// TIA Portal V21 export
// export: Created 2026-08-21T20:18:56.6399431Z, ExportSetting None, DisplayName Totally Integrated Automation Portal, DisplayVersion V21, DisplayName STEP 7 Professional, DisplayVersion V21, DisplayName STEP 7 Safety, DisplayVersion V21, DisplayName Tech WebApplication, DisplayVersion V21, DisplayName WinCC Basic/Comfort/Advanced, DisplayVersion V21, DisplayName WinCC Professional, DisplayVersion V21, DisplayName WinCC Unified, DisplayVersion V21
TYPE "UDT_Service_StepOrder"
   STRUCT
      stepNumber : Int := -1;   // actual number of step
      stepMonitoringTime : UDInt := 1000;   // step monitoring time
      parameter : "UDT_Service_IndexElement";   // start index of used parameters in parameter Array
   END_STRUCT;
END_TYPE
